FUNCTION_BLOCK FB_TemperaturOK_1
VAR_INPUT
	bEnable						:BOOL;			(* Enable FB signal *)
	bIn							:BOOL;			(* Temperature OK *)
	tTimeOutTempOK				:TIME := t#5s;		(* Temperature OK timeout *)
	tTimeOutTempNOK			:TIME := t#5s;		(* Temperature NOK timeout *)
END_VAR
VAR_OUTPUT
	bOut					:BOOL;			(* Temperature OK *)
	bError					:BOOL;			(* Error by temperature NOK *)
	udnErrorNo				:UDINT;
	udnMessageNo			:UDINT;
	sMsg					:STRING;
END_VAR
VAR
	bFirstTime			:BOOL;			(* First cycle *)
	tonDelayOK			:TON;			(* Temperatur delay ok *)
	tofWatchDog			:TOF;			(* Timer to off *)

END_VAR


IF NOT bFirstTime
THEN
	bError := FALSE;
	udnErrorNo := 0;
	udnMessageNo := 0;
	sMsg := '';
	tonDelayOK(
		IN := FALSE,
	          PT := tTimeOutTempOK
	);
	tofWatchDog(
		IN := FALSE,
	         PT := tTimeOutTempNOK
	);
	bFirstTime := TRUE;
END_IF;

(* Timer starts when came rising edge of signal *)
tonDelayOK(
	IN := bIn,
         PT := tTimeOutTempOK
);

tofWatchDog(
	IN := bIn,
         PT := tTimeOutTempNOK
);

IF tonDelayOK.Q
THEN
	bOut := TRUE;
    
ELSIF NOT tofWatchDog.Q
THEN
	bOut := FALSE;
    
END_IF;

END_FUNCTION_BLOCK

(* stored: Version 1.1.0.1, ProductVersion 3.1.4024.15
   POU FB_TemperaturOK_1: Id {3b054c07-6bba-4a4b-9667-edd75cc60ffe}, SpecialFunc None *)
